(* The principle is simple, a VRC should never open when B side pressure is greater than
the A side pressure. *)

FUNCTION F_VRC_DIODE_ILK : BOOL
VAR_INPUT

    i_stPGA : ST_VG; // A side pressure gauge
    i_stPGB	: ST_VG; // B side pressure gauge

END_VAR
VAR

    rHysterisis : REAL := 0;

    xInterlock: BOOL;
    rTolerance: REAL := 20;
END_VAR

(* The principle is simple, a VRC should never open when B side pressure is greater than the A side pressure. *)
rTolerance := 20;
F_VRC_DIODE_ILK := ((i_stPGA.rPRESS + rTolerance >= i_stPGB.rPRESS + rHysterisis) OR i_stPGA.xBAKEOUT) AND i_stPGA.xPRESS_OK AND i_stPGB.xPRESS_OK;

(* OK it gets a bit more complicated with hysterisis,

Now, if the F_VIC_DIODE_ILK is FALSE then some hysterisis is added to the B side. But if it's OK then we just stick with making sure that the A side is greater than the B side

*)
(*
IF NOT F_VIC_DIODE_ILK THEN
Hysterisis := 40;
ELSE
Hysterisis := 0;
END_IF
*)

END_FUNCTION

(* stored: Version 1.1.0.1
   POU F_VRC_DIODE_ILK: Id {0ea60bd7-e509-4e96-9cac-f7851bb32459}, SpecialFunc None *)
